Fanuc KAREL source: kb00195.KL

-- PROVISIONAL review KL for V940-1; original PC SHA256 ce4ae557cc6ef9f759a8313f8fd66a5cfc4b40a36376b92ec79fe280f3007ed5
-- Incomplete behavior may be omitted. Consult companion uncertainty JSON. Do not deploy.
PROGRAM KB00195
%NOLOCKGROUP
BEGIN
  -- V9_ZERO_TABLE_METADATA_HINT layout=0002_ascii; no indexed target words; source/name/runtime held
  -- UNRESOLVED_PC offsets 5-14; opcodes 3F,75
  -- UNRESOLVED_PC offsets 19-28; opcodes 3F,75
  -- UNRESOLVED_PC offsets 33-40; opcodes 9D,23
  -- UNRESOLVED_PC offsets 45-52; opcodes 9D,23
  -- UNRESOLVED_PC offsets 57-64; opcodes 9D,23
  -- UNRESOLVED_PC offsets 69-76; opcodes 9D,23
  -- UNRESOLVED_PC offsets 81-88; opcodes 9D,23
  -- UNRESOLVED_PC offsets 93-149; opcodes 27,22,2A,22,2A,22,22,22,22,22,22,31
  -- UNRESOLVED_PC offsets 154-158; opcodes 7F
END KB00195
